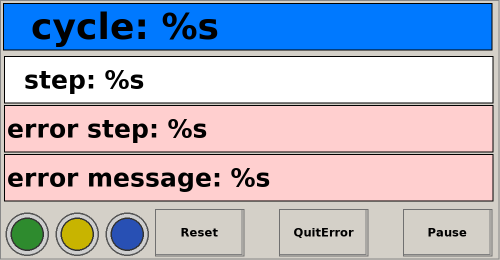
VISUALIZATION vis_Cycle_Control_1  // 500x260
VAR_IN_OUT
	fb: FB_SFC_Cycle;
END_VAR
VAR_INPUT
	sName: STRING:='Cycle name';
END_VAR
    Lamp1 (2,209 50x50), tooltip "Ready", variable: fb.bReady, style: Lamp-Lamp1-Green
    Lamp1 (102,209 50x50), tooltip "Done", variable: fb.bDone, style: Lamp-Lamp1-Blue
    Lamp1 (52,209 50x50), tooltip "Run", variable: fb.bRun, style: Lamp-Lamp1-Yellow
    RoundedRectangle (3,3 489x47), "cycle: %s", tooltip "POU name: %s", text variable: sName
        p4168582468: fb.refSFC.SFCErrorPOU
    RoundedRectangle (4,56 489x47), "step: %s", text variable: fb.refSFC.SFCCurrentStep, colour toggle: fb.ErrorSFC
    Button (155,209 89x47), "Reset"
        tap fb.bInit
    Button (403,209 89x47), "Pause", colour toggle: fb.refSFC.SFCPause
        toggle fb.refSFC.SFCPause
    Button (279,209 89x47), "QuitError", colour toggle: fb.ErrorSFC
        toggle fb.refSFC.SFCQuitError
    RoundedRectangle (4,105 489x47), "error step: %s", text variable: fb.sLastStepBefore_Error, colour toggle: fb.ErrorSFC
    RoundedRectangle (4,154 489x47), "error message: %s", text variable: fb.sError_Message, colour toggle: fb.ErrorSFC
END_VISUALIZATION

(* stored: Version 1.1.0.1, ProductVersion 3.1.4024.12
   Visu vis_Cycle_Control_1: Id {7989a24d-fb7d-432c-87e2-93c895632ed2} *)
